{ attribute 'Name':='TB_Prod-Test' }
{ attribute 'Timeout':='t#20s' }
{ attribute 'Owner':='TestOwner' }
{ attribute 'Category':='Math/multiplication and division ' }
FUNCTION_BLOCK FB_TestProd EXTENDS FB_TestCaseBase
VAR_INPUT
END_VAR
VAR_OUTPUT
END_VAR
VAR
	myFB : SampleLib.FB_Prod;   // instance of the function block to be tested
	expectedValue : UINT;       // value to be expected from this test
	result: UINT;				// calculated value, actual result of the function block call
END_VAR

// can of the function block to execute the test: 2 * 2 = 4
myFB(var1:= 2, var2:= 2, result=> result);

// Explicit assignment of the expected value, as the comparison is performed using the “any” data type
expectedValue:=4;

// Check the result against the expected value; if it does not match, the error message passed here is displayed
AssertEqual(anyActual:= result, anyExpected:= expectedValue, sMessage:= 'Multiplication with the FB_Prod function block is incorrect!');

// in the event that the result of the comparison matches, confirmation that the test case was successful and that no further tests will be carried out in this function block
Succeed();

//Must be implemented if you want to use fastmode
METHOD CleanUp : BOOL
CleanUp:=true;
END_METHOD

END_FUNCTION_BLOCK

(* stored: Version 1.1.0.1, ProductVersion 3.1.4026.21
   POU FB_TestProd: Id {e2a37850-0368-4db9-a7a1-9065adaee9ca}, SpecialFunc None
   Method CleanUp: Id {dbc2c251-0820-4004-9560-f1549cb1fb1f} *)
